(* IEC 61131-3 sources: 2026_Projet_YGO_ExcavatriceDragage/TOOLS/TEST_AUTO_CI/RESULTS/L_SIMULATION/tests (part 3) *)

(* ---- test_fb_sim_position_sensor.st ---- *)
(* T300 - Tests unitaires du capteur cumulatif M3. *)
TEST 'TC-T300-SEN-010 Hysteresis cumulative conserve le mot thermometre'
VAR
    fb : FB_Sim_PositionSensor;
END_VAR
    fb.Enable := TRUE;
    fb.Threshold_M := 5.0;
    fb.Hysteresis_M := 0.02;
    fb.Position_M := 4.99;
    fb();
    ASSERT_TRUE(fb.ElectricalOutput, 'Position sous seuil active DI cumulative');
    fb.Position_M := 5.01;
    fb();
    ASSERT_TRUE(fb.ElectricalOutput, 'Hysteresis maintient DI dans la bande');
    fb.Position_M := 5.03;
    fb();
    ASSERT_FALSE(fb.ElectricalOutput, 'Sortie au-dessus de seuil+hysteresis');
    fb.Position_M := 4.99;
    fb();
    ASSERT_FALSE(fb.ElectricalOutput, 'Retour dans bande ne re-declenche pas');
    fb.Position_M := 4.97;
    fb();
    ASSERT_TRUE(fb.ElectricalOutput, 'Retour sous seuil-hysteresis re-declenche');
END_TEST

TEST 'TC-T300-SEN-030 Episode intermittent est borne et rejoint la position'
VAR
    fb : FB_Sim_PositionSensor;
    i : INT;
END_VAR
    fb.Enable := TRUE;
    fb.Threshold_M := 5.0;
    fb.Position_M := 4.0;
    fb.IntermittenceActive := TRUE;
    fb.IntermittenceDurationS := 1.0;
    fb.IntermittencePeriodS := 0.12;
    fb.CycleTimeS := 0.01;
    fb();
    fb.Position_M := 6.0;
    FOR i := 1 TO 120 DO
        fb();
    END_FOR;
    ASSERT_FALSE(fb.EpisodeActive, 'Episode termine avant 1.2 s');
    ASSERT_FALSE(fb.ElectricalOutput, 'DI rejoint l etat mecanique final');
    ASSERT_GT(fb.TransitionCount, 2, 'Pertes/reprises publiees, sans front permanent');
END_TEST

TEST 'TC-T300-SEN-031 Recroisements mecaniques ne reinitialisent pas episode'
VAR
    fb : FB_Sim_PositionSensor;
    i : INT;
END_VAR
    fb.Enable := TRUE;
    fb.Threshold_M := 5.0;
    fb.Position_M := 4.0;
    fb.IntermittenceActive := TRUE;
    fb.IntermittenceDurationS := 1.0;
    fb.IntermittencePeriodS := 0.12;
    fb.CycleTimeS := 0.01;
    fb();
    FOR i := 1 TO 40 DO
        IF (i MOD 2) = 0 THEN
            fb.Position_M := 4.0;
        ELSE
            fb.Position_M := 6.0;
        END_IF;
        fb();
    END_FOR;
    fb.Position_M := 6.0;
    FOR i := 1 TO 70 DO
        fb();
    END_FOR;
    ASSERT_FALSE(fb.EpisodeActive, 'Recroisements ne prolongent pas episode au-dela de 1 s');
    ASSERT_FALSE(fb.ElectricalOutput, 'Etat final suit dernier franchissement mecanique');
END_TEST

TEST 'TC-T300-SEN-040 Cent graines deterministes bornent la stabilisation'
VAR
    fb : FB_Sim_PositionSensor;
    i : INT;
    j : INT;
END_VAR
    FOR i := 1 TO 100 DO
        fb.Enable := FALSE;
        fb();
        fb.Enable := TRUE;
        fb.Threshold_M := 5.0;
        fb.Position_M := 4.0;
        fb.IntermittenceActive := TRUE;
        fb.IntermittenceDurationS := 1.0;
        fb.IntermittencePeriodS := 0.12;
        fb.CycleTimeS := 0.01;
        fb.ScenarioSeed := DINT_TO_UDINT(i);
        fb();
        fb.Position_M := 6.0;
        FOR j := 1 TO 120 DO
            fb();
        END_FOR;
        ASSERT_FALSE(fb.EpisodeActive, 'Chaque graine termine son episode avant 1.2 s');
        ASSERT_FALSE(fb.ElectricalOutput, 'Chaque graine rejoint la position finale');
        ASSERT_GE(fb.EpisodeTogglePeriodS, 0.084, 'Periode aleatoire >= 70 % nominal');
        ASSERT_LE(fb.EpisodeTogglePeriodS, 0.156, 'Periode aleatoire <= 130 % nominal');
    END_FOR;
END_TEST

(* T300 P-A / C1-C2 — profil « BLIP COURT » : excursions electriques courtes, parametrables,
   independantes du train ~1 s ci-dessus. Signatures de la trace terrain du 2026-09-04 :
   Tremie contradictoire pendant 2 echantillons a 12,24 s ; PV reactive 1 echantillon a 14,94 s.
   Grille de test = 100 ms, celle de la trace. *)
TEST 'TC-T300-SEN-050 Blip court : largeur parametrable, deux sens, profil 1 s intact'
VAR
    fb : FB_Sim_PositionSensor;
    i : INT;
    excursions : INT;
    baseCount : UDINT;
END_VAR
    (* ---- (1) Sortie de zone, excursion 0,1 s => 1 echantillon (signature PV) ---- *)
    fb.Enable := TRUE;
    fb.Threshold_M := 5.0;
    fb.Hysteresis_M := 0.02;
    fb.CycleTimeS := 0.1;
    fb.ElectricalDelayS := 0.0;
    fb.Position_M := 4.0;
    fb();
    ASSERT_TRUE(fb.ElectricalOutput, 'Depart : dans la zone capteur');
    baseCount := fb.TransitionCount;
    fb.BlipTransitions := 1;
    fb.BlipDurationS := 0.1;
    fb.Position_M := 6.0;
    fb();
    excursions := 0;
    FOR i := 1 TO 6 DO
        fb();
        IF fb.ElectricalOutput <> fb.RawDetected THEN
            excursions := excursions + 1;
        END_IF;
    END_FOR;
    ASSERT_EQ(excursions, 1, 'Blip 0,1 s a 100 ms = 1 echantillon contradictoire');
    ASSERT_EQ(fb.TransitionCount - baseCount, 3, '1 front nominal + 2 fronts du blip');
    ASSERT_FALSE(fb.BlipActive, 'Blip borne et termine');
    ASSERT_FALSE(fb.ElectricalOutput, 'Sortie rendue a l etat mecanique final');

    (* ---- (2) Meme sens, excursion 0,2 s => 2 echantillons (signature Tremie) ---- *)
    fb.Enable := FALSE;
    fb();
    fb.Enable := TRUE;
    fb.BlipTransitions := 1;
    fb.BlipDurationS := 0.2;
    fb.Position_M := 4.0;
    fb();
    fb.Position_M := 6.0;
    fb();
    excursions := 0;
    FOR i := 1 TO 8 DO
        fb();
        IF fb.ElectricalOutput <> fb.RawDetected THEN
            excursions := excursions + 1;
        END_IF;
    END_FOR;
    ASSERT_EQ(excursions, 2, 'Blip 0,2 s a 100 ms = 2 echantillons contradictoires');
    ASSERT_FALSE(fb.ElectricalOutput, 'Sortie rendue a l etat mecanique final');

    (* ---- (3) Sens INVERSE : entree en zone (front montant) — symetrie AC5 ---- *)
    fb.Enable := FALSE;
    fb();
    fb.Enable := TRUE;
    fb.BlipTransitions := 1;
    fb.BlipDurationS := 0.2;
    fb.Position_M := 6.0;
    fb();
    ASSERT_FALSE(fb.ElectricalOutput, 'Depart : hors zone capteur');
    fb.Position_M := 4.0;
    fb();
    excursions := 0;
    FOR i := 1 TO 8 DO
        fb();
        IF fb.ElectricalOutput <> fb.RawDetected THEN
            excursions := excursions + 1;
        END_IF;
    END_FOR;
    ASSERT_EQ(excursions, 2, 'Symetrie : excursion equivalente a l entree en zone');
    ASSERT_TRUE(fb.ElectricalOutput, 'Sortie rendue a l etat mecanique final (dans la zone)');

    (* ---- (4) Blip DESACTIVE : le profil historique reste strictement inchange ---- *)
    fb.Enable := FALSE;
    fb();
    fb.Enable := TRUE;
    fb.BlipTransitions := 0;
    fb.Position_M := 4.0;
    fb();
    baseCount := fb.TransitionCount;
    fb.Position_M := 6.0;
    fb();
    excursions := 0;
    FOR i := 1 TO 10 DO
        fb();
        IF fb.ElectricalOutput <> fb.RawDetected THEN
            excursions := excursions + 1;
        END_IF;
    END_FOR;
    ASSERT_EQ(excursions, 0, 'Blip desactive : aucune excursion inventee');
    ASSERT_EQ(fb.TransitionCount - baseCount, 1, 'Blip desactive : seul le front nominal');
END_TEST

(* ---- test_fb_sim_safety.st ---- *)
(* =======================================================================
   Automated Unit Test - FB_Sim_Safety
   ======================================================================= *)
TEST 'TC-P13-SAF-001 Enable FALSE -> boucle AU ouverte'
VAR
    fb : FB_Sim_Safety;
END_VAR
    fb.Enable := FALSE;
    fb.SimChainOkBit := TRUE;
    fb();
    ASSERT_FALSE(fb.SimChainOk, 'Enable FALSE -> SimChainOk FALSE');
    ASSERT_FALSE(fb.SimContactorOk, 'Enable FALSE -> SimContactorOk FALSE');
END_TEST

TEST 'TC-P13-SAF-002 Pilotage boucle AU saine par SimChainOkBit et armement contacteur'
VAR
    fb : FB_Sim_Safety;
END_VAR
    fb.Enable := TRUE;
    fb.SimChainOkBit := TRUE; (* Chaine AU fermee par operateur *)
    fb();

    (* Ecoulement tempo de fermeture chaine (50ms = 60ms avancee) *)
    ADVANCE_TIME(60000000);
    fb();
    ASSERT_TRUE(fb.SimChainOk, 'SimChainOkBit TRUE -> SimChainOk TRUE apres tempo relais');

    (* Impulsion armement tenue 100ms (temps de collage contacteur) *)
    ADVANCE_TIME(10000000);
    fb.EmergencyArming := TRUE;
    fb();
    ADVANCE_TIME(110000000);
    fb();
    ASSERT_TRUE(fb.SimContactorOk, 'EmergencyArming soutenu -> SimContactorOk TRUE (engage)');

    (* Relachement impulsion -> auto-maintien *)
    ADVANCE_TIME(10000000);
    fb.EmergencyArming := FALSE;
    fb();
    ASSERT_TRUE(fb.SimContactorOk, 'Fin pulse -> Auto-maintien contacteur maintenu');
END_TEST

TEST 'TC-T306-SAF-003 Injection defaut rotation de phases par SimPhaseRotationOkBit'
VAR
    fb : FB_Sim_Safety;
END_VAR
    (* Phases saines : SimPhaseRotationOkBit=TRUE -> sortie TRUE (aucun defaut) *)
    fb.Enable := TRUE;
    fb.SimPhaseRotationOkBit := TRUE;
    fb();
    ASSERT_TRUE(fb.SimPhaseRotationOk, 'SimPhaseRotationOkBit TRUE -> SimPhaseRotationOk TRUE (phases saines)');

    (* Defaut injecte : SimPhaseRotationOkBit=FALSE -> sortie FALSE (PhaseRotationOk_DI tombe) *)
    fb.SimPhaseRotationOkBit := FALSE;
    fb();
    ASSERT_FALSE(fb.SimPhaseRotationOk, 'SimPhaseRotationOkBit FALSE -> SimPhaseRotationOk FALSE (defaut rotation de phases)');

    (* Retour a sain : nouveau passage a TRUE -> sortie TRUE *)
    fb.SimPhaseRotationOkBit := TRUE;
    fb();
    ASSERT_TRUE(fb.SimPhaseRotationOk, 'SimPhaseRotationOkBit TRUE apres FALSE -> SimPhaseRotationOk TRUE');
END_TEST

(* ---- test_fb_sim_suspended_load.st ---- *)
TEST 'TC-T300-MEC-010 Charge au repos ne cree pas d energie'
VAR
    fb : FB_Sim_SuspendedLoad;
    i : INT;
END_VAR
    fb.Enable := TRUE;
    fb.CycleTime_S := 0.01;
    FOR i := 1 TO 6000 DO
        fb();
    END_FOR;
    ASSERT_EQ(fb.Angle_Rad, 0.0, 'Angle nul sans excitation pendant 60 s');
    ASSERT_EQ(fb.AngularVelocity_RadPerS, 0.0, 'Vitesse angulaire nulle sans excitation');
END_TEST

TEST 'TC-T300-MEC-040 Acceleration excite charge et reaction reste conditionnee au frein'
VAR
    fb : FB_Sim_SuspendedLoad;
    i : INT;
END_VAR
    fb.Enable := TRUE;
    fb.CartAcceleration_Mps2 := 1.0;
    fb.BrakeMechanicallyOpen := FALSE;
    fb.CycleTime_S := 0.01;
    fb();
    ASSERT_TRUE(ABS(fb.Angle_Rad) > 0.0, 'Acceleration excite le pendule');
    ASSERT_EQ(fb.VelocityReaction_Mps, 0.0, 'Frein serre bloque reaction chariot');
    fb.BrakeMechanicallyOpen := TRUE;
    fb.CartAcceleration_Mps2 := 0.0;
    FOR i := 1 TO 10 DO
        fb();
    END_FOR;
    ASSERT_TRUE(ABS(fb.VelocityReaction_Mps) > 0.0, 'Frein ouvert publie reaction charge');
END_TEST

TEST 'TC-T300-MEC-020 Convergence pendule entre pas 10 ms et 5 ms'
VAR
    fb10 : FB_Sim_SuspendedLoad;
    fb5 : FB_Sim_SuspendedLoad;
    i : INT;
END_VAR
    fb10.Enable := TRUE;
    fb10.BrakeMechanicallyOpen := TRUE;
    fb10.CartAcceleration_Mps2 := 1.0;
    fb10.CycleTime_S := 0.01;
    fb5.Enable := TRUE;
    fb5.BrakeMechanicallyOpen := TRUE;
    fb5.CartAcceleration_Mps2 := 1.0;
    fb5.CycleTime_S := 0.005;
    fb10();
    fb5();
    fb5();
    fb10.CartAcceleration_Mps2 := 0.0;
    fb5.CartAcceleration_Mps2 := 0.0;
    FOR i := 1 TO 100 DO
        fb10();
        fb5();
        fb5();
    END_FOR;
    ASSERT_LT(ABS(fb10.Angle_Rad - fb5.Angle_Rad), 0.01,
        'Ecart angle inferieur a 10 mrad apres 1 s');
    ASSERT_LT(ABS(fb10.VelocityReaction_Mps - fb5.VelocityReaction_Mps), 0.001,
        'Ecart reaction inferieur a 1 mm/s apres 1 s');
END_TEST

(* ---- test_fb_sim_translation.st ---- *)
(* T300 - Tests du modele dynamique M3. *)
TEST 'TC-T300-TR-001 Etat sur desactive est P1 sans mouvement'
VAR
    fb : FB_Sim_Translation;
END_VAR
    fb.Enable := FALSE;
    fb();
    ASSERT_FALSE(fb.PosTremie, 'P1 ne doit pas annoncer Tremie');
    ASSERT_TRUE(fb.PosP1, 'Etat de repli deterministe sur P1');
    ASSERT_TRUE(fb.PosMaintenance, 'Mot thermometre P1 attendu');
    ASSERT_EQ(fb.ActualFrequency_Hz, 0.0, 'Frequence nulle');
    ASSERT_FALSE(fb.BrakeContactOpen, 'Frein ferme');
END_TEST

(* T301/L1 -- the isolated model receives geometry and gain.  The static G518
   check proves the PRG_02 -> SimBench wiring; these cases prove that those
   inputs are actually consumed by the simulated plant. *)
TEST 'TC-T301-SRC-001 Position P1 recue initialise le chariot sans geometrie locale'
VAR
    fb : FB_Sim_Translation;
END_VAR
    fb.PosTremie_M := 2.0;
    fb.PosPV_M := 3.0;
    fb.PosP2_M := 5.0;
    fb.PosP1_M := 7.0;
    fb.PosMaintenance_M := 11.0;
    fb.Enable := FALSE;
    fb();
    ASSERT_NEAR(fb.PositionTrue_M, 7.0, 0.0001,
        'Repli positionne le chariot sur PosP1_M recu');
    ASSERT_TRUE(fb.PosP1, 'Repli publie P1 apres initialisation sur la position recue');
END_TEST

TEST 'TC-T301-SRC-002 Gain recu convertit la frequence retournee en vitesse'
VAR
    fb : FB_Sim_Translation;
    i : INT;
END_VAR
    fb.PosTremie_M := 0.0;
    fb.PosPV_M := 10.0;
    fb.PosP2_M := 20.0;
    fb.PosP1_M := 30.0;
    fb.PosMaintenance_M := 40.0;
    fb.GainMetersPerHzSec := 0.03;
    fb.MaxFreq_Hz := 20.0;
    fb.Enable := FALSE;
    fb();
    fb.Enable := TRUE;
    fb.ReqTremie := TRUE;
    fb.SpeedTgt_Pct := 100.0;
    fb.BrakeReleaseCmd := TRUE;
    fb.BrakeOpenDelayS := 0.0;
    fb.LoadReactionGain_Mps2 := 0.0;
    FOR i := 1 TO 400 DO
        fb();
    END_FOR;
    ASSERT_NEAR(fb.ActualFrequency_Hz, 20.0, 0.05,
        'Frequence maximale recue appliquee');
    ASSERT_NEAR(fb.VelocityTrue_Mps, -0.6, 0.02,
        'Vitesse = sens x gain recu x frequence retournee');
END_TEST

TEST 'TC-T300-SEN-010 Les deux extremites publient les mots thermometres valides'
VAR
    fb : FB_Sim_Translation;
    i : INT;
END_VAR
    fb.Enable := FALSE;
    fb();
    fb.Enable := TRUE;
    fb.ReqTremie := TRUE;
    fb.SpeedTgt_Pct := 100.0;
    fb.BrakeReleaseCmd := TRUE;
    fb.BrakeOpenDelayS := 0.0;
    fb.FullTravelTimeS := 0.5;
    fb.SensorElectricalDelayS := 0.0;
    FOR i := 1 TO 400 DO
        fb();
    END_FOR;
    ASSERT_TRUE(fb.PosTremie, 'Tremie active a la butee 0 m');
    ASSERT_TRUE(fb.PosPV, 'PV cumulatif actif a Tremie');
    ASSERT_TRUE(fb.PosP2, 'P2 cumulatif actif a Tremie');
    ASSERT_TRUE(fb.PosP1, 'P1 cumulatif actif a Tremie');
    ASSERT_TRUE(fb.PosMaintenance, 'Maintenance cumulatif actif a Tremie');
    ASSERT_EQ(fb.VelocityTrue_Mps, 0.0, 'Butee Tremie absorbe la vitesse chariot');

    fb.Enable := FALSE;
    fb();
    fb.Enable := TRUE;
    fb.ReqTremie := FALSE;
    fb.ReqMaintenance := TRUE;
    fb.SpeedTgt_Pct := 100.0;
    fb.BrakeReleaseCmd := TRUE;
    fb.BrakeOpenDelayS := 0.0;
    fb.FullTravelTimeS := 0.5;
    fb.SensorElectricalDelayS := 0.0;
    FOR i := 1 TO 400 DO
        fb();
    END_FOR;
    ASSERT_FALSE(fb.PosTremie, 'Tremie inactif a Maintenance');
    ASSERT_FALSE(fb.PosPV, 'PV inactif a Maintenance');
    ASSERT_FALSE(fb.PosP2, 'P2 inactif a Maintenance');
    ASSERT_FALSE(fb.PosP1, 'P1 inactif a Maintenance');
    ASSERT_FALSE(fb.PosMaintenance, 'Maintenance inactif a la butee pour mot 00000');
    ASSERT_EQ(fb.VelocityTrue_Mps, 0.0, 'Butee Maintenance absorbe la vitesse chariot');
END_TEST

TEST 'TC-T300-SEN-011 Le capteur PV commute au franchissement vers Tremie'
VAR
    fb : FB_Sim_Translation;
    i : INT;
    pvWasFalse : BOOL;
    pvTurnedTrue : BOOL;
END_VAR
    fb.Enable := TRUE;
    fb.ReqTremie := TRUE;
    fb.SpeedTgt_Pct := 100.0;
    fb.BrakeReleaseCmd := TRUE;
    fb.FullTravelTimeS := 8.0;
    fb.SensorElectricalDelayS := 0.0;
    pvWasFalse := FALSE;
    pvTurnedTrue := FALSE;
    FOR i := 1 TO 700 DO
        fb();
        IF NOT fb.PosPV THEN
            pvWasFalse := TRUE;
        END_IF;
        IF pvWasFalse AND fb.PosPV THEN
            pvTurnedTrue := TRUE;
        END_IF;
    END_FOR;
    ASSERT_TRUE(pvWasFalse, 'PV initialement inactif a P1');
    ASSERT_TRUE(pvTurnedTrue, 'PV actif apres franchissement vers Tremie');
END_TEST

TEST 'TC-T300-DRV-020 Rampe terrain 20 Hz par seconde'
VAR
    fb : FB_Sim_Translation;
    i : INT;
END_VAR
    fb.Enable := TRUE;
    fb.ReqTremie := TRUE;
    fb.SpeedTgt_Pct := 0.0;
    fb.BrakeReleaseCmd := TRUE;
    fb();
    fb.SpeedTgt_Pct := 100.0;
    FOR i := 1 TO 100 DO
        fb();
    END_FOR;
    ASSERT_GT(fb.FrequencyCmd_Hz, 19.7, 'Rampe apres 1 s >= 19.7 Hz');
    ASSERT_LT(fb.FrequencyCmd_Hz, 20.3, 'Rampe apres 1 s <= 20.3 Hz');
    ASSERT_LT(fb.ActualFrequency_Hz, fb.FrequencyCmd_Hz, 'Retour dynamique derriere la consigne');
    ASSERT_GT(fb.ActualFrequency_Hz, 16.0, 'Retour coherent avec tau 150 ms');
END_TEST

TEST 'TC-T300-BRK-025 Frein temporise et retour distinct'
VAR
    fb : FB_Sim_Translation;
    i : INT;
END_VAR
    fb.Enable := TRUE;
    fb.BrakeReleaseCmd := TRUE;
    fb.BrakeOpenDelayS := 0.10;
    fb();
    ASSERT_TRUE(fb.BrakeCoilEnergized, 'Bobine active immediatement sur ordre');
    FOR i := 1 TO 8 DO
        fb();
    END_FOR;
    ASSERT_FALSE(fb.BrakeContactOpen, 'Pas de confirmation avant 90 ms');
    fb();
    fb();
    ASSERT_TRUE(fb.BrakeMechanicallyOpen, 'Ouverture mecanique apres delai');
    ASSERT_TRUE(fb.BrakeContactOpen, 'Retour auxiliaire apres delai');
END_TEST

TEST 'TC-T300-MEC-010 Le chariot suit la frequence et excite la charge'
VAR
    fb : FB_Sim_Translation;
    i : INT;
    startPosition_M : REAL;
END_VAR
    fb.Enable := TRUE;
    fb.ReqTremie := TRUE;
    fb.SpeedTgt_Pct := 100.0;
    fb.BrakeReleaseCmd := TRUE;
    fb.BrakeOpenDelayS := 0.0;
    fb();
    startPosition_M := fb.PositionTrue_M;
    FOR i := 1 TO 100 DO
        fb();
    END_FOR;
    ASSERT_LT(fb.PositionTrue_M, startPosition_M, 'Deplacement reel vers Tremie');
    ASSERT_LT(fb.VelocityTrue_Mps, 0.0, 'Vitesse signee vers Tremie');
    ASSERT_TRUE(ABS(fb.LoadAngle_Rad) > 0.0001, 'Acceleration excite le pendule');
END_TEST

TEST 'TC-T300-MEC-030 Commandes contradictoires restent neutres'
VAR
    fb : FB_Sim_Translation;
    i : INT;
    startPosition_M : REAL;
END_VAR
    fb.Enable := TRUE;
    fb.ReqTremie := TRUE;
    fb.ReqMaintenance := TRUE;
    fb.SpeedTgt_Pct := 100.0;
    fb.BrakeReleaseCmd := TRUE;
    fb.BrakeOpenDelayS := 0.0;
    fb();
    startPosition_M := fb.PositionTrue_M;
    FOR i := 1 TO 50 DO
        fb();
    END_FOR;
    ASSERT_EQ(fb.FrequencyCmd_Hz, 0.0, 'Aucune excitation avec deux sens');
    ASSERT_EQ(fb.PositionTrue_M, startPosition_M, 'Position conservee');
END_TEST

TEST 'TC-T300-SEN-030 Episode capteur intermittent rejouable avant stabilisation'
VAR
    fb : FB_Sim_Translation;
    i : INT;
END_VAR
    fb.Enable := TRUE;
    fb.ReqMaintenance := TRUE;
    fb.SpeedTgt_Pct := 0.0;
    fb.BrakeReleaseCmd := TRUE;
    fb.BrakeOpenDelayS := 0.0;
    fb.FullTravelTimeS := 0.5;
    fb.SensorStabilizationS := 1.0;
    fb.SensorIntermittenceActive := TRUE;
    fb.SensorLoadAngleTriggerRad := 0.0;
    fb.SensorIntermittencePeriodS := 0.12;
    fb();
    fb.SpeedTgt_Pct := 100.0;
    FOR i := 1 TO 250 DO
        fb();
    END_FOR;
    ASSERT_GT(fb.SensorTransitionCount, 1, 'Au moins deux fronts DI sont publies pendant episode');
    ASSERT_FALSE(fb.PosP1, 'DI rejoint la position mecanique apres episode');
END_TEST

TEST 'TC-T300-CAM-100 Matrice 48 scenarios par 100 graines respecte invariants'
VAR
    fb : FB_Sim_Translation;
    direction : INT;
    loadProfile : INT;
    regime : INT;
    perturbation : INT;
    seed : INT;
    i : INT;
END_VAR
    FOR direction := 1 TO 2 DO
        FOR loadProfile := 1 TO 2 DO
            FOR regime := 1 TO 3 DO
                FOR perturbation := 1 TO 4 DO
                    FOR seed := 1 TO 100 DO
                        fb.Enable := FALSE;
                        fb();
                        fb.Enable := TRUE;
                        fb.ReqTremie := direction = 1;
                        fb.ReqMaintenance := direction = 2;
                        fb.SpeedTgt_Pct := 100.0;
                        fb.BrakeReleaseCmd := TRUE;
                        fb.FullTravelTimeS := 0.5;
                        fb.SensorElectricalDelayS := 0.0;
                        fb.SensorScenarioSeed := DINT_TO_UDINT(seed);
                        fb.SensorIntermittenceActive := perturbation = 3;
                        fb.SensorLoadAngleTriggerRad := 0.0;
                        IF loadProfile = 1 THEN
                            fb.LoadReactionGain_Mps2 := 0.0;
                        ELSE
                            fb.LoadReactionGain_Mps2 := 0.20;
                        END_IF;
                        IF perturbation = 4 THEN
                            fb.BrakeOpenDelayS := 0.30;
                        ELSE
                            fb.BrakeOpenDelayS := 0.0;
                        END_IF;
                        fb();
                        FOR i := 1 TO 200 DO
                            IF (regime = 2) AND (i = 80) THEN
                                fb.SpeedTgt_Pct := 0.0;
                            ELSIF (regime = 3) AND (i = 80) THEN
                                fb.SpeedTgt_Pct := 0.0;
                                fb.BrakeReleaseCmd := FALSE;
                            END_IF;
                            fb();
                            ASSERT_GE(fb.PositionTrue_M, 0.0, 'Course mecanique jamais inferieure a Tremie');
                            ASSERT_LE(fb.PositionTrue_M, 30.0, 'Course mecanique jamais superieure a Maintenance');
                            ASSERT_GE(fb.ActualFrequency_Hz, 0.0, 'Retour variateur non negatif');
                            ASSERT_LE(fb.ActualFrequency_Hz, 50.0, 'Retour variateur borne a 50 Hz');
                            IF perturbation <> 3 THEN
                                ASSERT_TRUE((NOT fb.PosTremie) OR fb.PosPV,
                                    'Mot thermometre : Tremie implique PV');
                                ASSERT_TRUE((NOT fb.PosPV) OR fb.PosP2,
                                    'Mot thermometre : PV implique P2');
                                ASSERT_TRUE((NOT fb.PosP2) OR fb.PosP1,
                                    'Mot thermometre : P2 implique P1');
                                ASSERT_TRUE((NOT fb.PosP1) OR fb.PosMaintenance,
                                    'Mot thermometre : P1 implique Maintenance');
                            END_IF;
                        END_FOR;
                    END_FOR;
                END_FOR;
            END_FOR;
        END_FOR;
    END_FOR;
END_TEST

(* T300 P-A / C4 — traversee de la faute frein dans le composite : prouve que l'entree
   descend jusqu'a FB_Sim_TranslationBrake et que la sortie remonte, sans toucher au
   nominal (premier palier d'assertions). *)
TEST 'TC-T300-BRK-041 Faute frein traverse le composite M3 (fermeture en mouvement)'
VAR
    fb : FB_Sim_Translation;
    i : INT;
END_VAR
    fb.Enable := TRUE;
    fb.ReqMaintenance := TRUE;
    fb.SpeedTgt_Pct := 100.0;
    fb.BrakeReleaseCmd := TRUE;
    fb.BrakeOpenDelayS := 0.0;
    fb();
    ASSERT_TRUE(fb.BrakeMechanicallyOpen, 'Frein ouvert au depart');
    FOR i := 1 TO 200 DO
        fb();
    END_FOR;
    ASSERT_GT(fb.ActualFrequency_Hz, 0.5, 'Chariot en mouvement (frequence non nulle)');
    ASSERT_TRUE(fb.BrakeMechanicallyOpen, 'NOMINAL : frein ouvert tant que la vitesse est non nulle');
    ASSERT_FALSE(fb.BrakeFaultCloseActive, 'Aucune faute par defaut');

    fb.BrakeFaultCloseWhileRunning := TRUE;
    FOR i := 1 TO 12 DO
        fb();
    END_FOR;
    ASSERT_TRUE(fb.BrakeFaultCloseActive, 'Faute frein relayee par le composite');
    ASSERT_GT(fb.ActualFrequency_Hz, 0.5, 'Vitesse encore non nulle a la fermeture');
    ASSERT_FALSE(fb.BrakeMechanicallyOpen, 'Faute : frein mecaniquement serre en mouvement');
END_TEST

(* T300 P-A / C3 — deceleration libre. Trace terrain 2026-09-04 : commande retiree a
   14,67 s alors que 33,98 Hz etaient retournes ; le chariot a continue d'avancer pendant
   1,49 s jusqu'a l'arret a 16,16 s. La distance de roue libre correspondante est une
   ESTIMATION (la trace ne contient aucune variable de position) : ordre de grandeur
   1,1 a 1,3 m selon la methode d'integration, jamais parcourus par le modele avant ce
   correctif qui annulait la vitesse au scan de retrait de commande.
   Le pas FullTravelTimeS est allonge (60 s) pour que le scenario reste loin des butees
   mecaniques et que l'oracle porte sur la SEULE deceleration libre, pas sur un choc. *)
TEST 'TC-T300-DRV-070 Deceleration libre : le chariot avance encore apres retrait de commande'
VAR
    fb : FB_Sim_Translation;
    i : INT;
    posAtCut_M : REAL;
END_VAR
    fb.Enable := TRUE;
    fb.ReqMaintenance := TRUE;
    fb.SpeedTgt_Pct := 100.0;
    fb.BrakeReleaseCmd := TRUE;
    fb.BrakeOpenDelayS := 0.0;
    (* Echelle par defaut du banc : palier 50 Hz (maximum variateur), 0,02 m/(Hz.s), rampe d'arret 25 Hz/s. *)
    (* Charge neutralisee : l'oracle porte sur la SEULE deceleration libre du variateur.
       Sans cela, le droop de charge (0,5 Hz par rad/s) peut faire passer ActualFrequency
       sous 39,5 Hz et rendre l'assertion de palier marginale — bruit, pas verite. *)
    fb.LoadFrequencyDroopGain_Hz := 0.0;
    fb.LoadReactionGain_Mps2 := 0.0;
    FOR i := 1 TO 400 DO
        fb();
    END_FOR;
    ASSERT_NEAR(fb.ActualFrequency_Hz, 50.0, 0.5, 'Palier 50 Hz etabli avant le retrait');
    ASSERT_LT(fb.PositionTrue_M, 30.0, 'Chariot encore hors butee (scenario non pollue)');

    (* Retrait total de la commande : plus aucune requete, consigne a zero. *)
    fb.ReqMaintenance := FALSE;
    fb.ReqTremie := FALSE;
    fb.SpeedTgt_Pct := 0.0;
    fb();
    ASSERT_GT(fb.ActualFrequency_Hz, 0.5, 'Le variateur retourne encore de la vitesse au retrait');
    posAtCut_M := fb.PositionTrue_M;

    (* Roue libre : la position doit continuer de varier tant que ActualFrequency_Hz > 0.
       Seuil = borne BASSE de la bande de reference trace (R2-O9 : 0,9 a 1,3 m). Le modele
       parcourt davantage (~2,2 m) car sa rampe de descente dure 2,0 s contre 1,49 s mesures :
       ecart de fidelite ASSUME, borne haute verifiee separement. Avant correctif : ~0,1 m. *)
    FOR i := 1 TO 300 DO
        fb();
    END_FOR;
    ASSERT_NEAR(fb.ActualFrequency_Hz, 0.0, 0.01, 'Retour variateur revenu a zero');
    ASSERT_GE(fb.PositionTrue_M - posAtCut_M, 0.9,
        'Roue libre >= borne basse trace (avant correctif : ~0,1 m)');
    ASSERT_LE(fb.PositionTrue_M - posAtCut_M, 3.0, 'Roue libre bornee (pas d emballement)');
    ASSERT_LE(fb.PositionTrue_M, 30.0, 'Course mecanique respectee');
END_TEST

(* T300 P-A / C5 — perte DEFINITIVE du capteur Tremie apres arret serre.
   Trace terrain 2026-09-04 : a 26,437 s le chariot entre en zone Tremie pendant que la
   commande est retiree ; le capteur retombe a 26,537 s et n'est JAMAIS repris sur les
   8,6 s restantes (PLAN_T300 §38 : perte unique post-arret, pas une oscillation entretenue).
   EndStopRecoilMax_M = 0 conserve le comportement historique (position ET vitesse figees,
   decision de review tracee) : les deux regimes sont verifies ici. *)
TEST 'TC-T300-SEN-052 Recul borne a la butee Tremie : DI perdue PUIS reprise oscillante (ecart trace)'
VAR
    fb : FB_Sim_Translation;
    i : INT;
    scansToFall : INT;
    scansActive : INT;
END_VAR
    (* --- (0) NON-REGRESSION : recul non autorise => comportement historique inchange --- *)
    fb.Enable := TRUE;
    fb.ReqTremie := TRUE;
    fb.SpeedTgt_Pct := 100.0;
    fb.BrakeReleaseCmd := TRUE;
    fb.BrakeOpenDelayS := 0.0;
    fb.SensorElectricalDelayS := 0.0;
    fb.EndStopRecoilMax_M := 0.0;
    (* T361 — pas de temps PINCE ici : l'oracle de ce cas est le recul a la butee, pas
       l'echelle odometrique. Le scenario vient de la trace du 2026-09-04 (quelques
       secondes de trajet) et le defaut du FB est passe de 8,0 s a 37,5 s pour s'aligner
       sur le gain reel : sans ce pas explicite, 900 scans (9 s) ne suffiraient plus a
       atteindre la butee Tremie depuis 20 m et le cas testerait autre chose que son objet. *)
    fb.FullTravelTimeS := 8.0;
    FOR i := 1 TO 900 DO
        fb();
    END_FOR;
    ASSERT_TRUE(fb.PosTremie, 'Historique : DI Tremie TENUE a la butee quand le recul est interdit');
    ASSERT_NEAR(fb.PositionTrue_M, 0.0, 0.001, 'Historique : position figee a la butee');

    (* --- (1) Recul borne autorise : la charge ressort le chariot de la zone --- *)
    fb.Enable := FALSE;
    fb();
    fb.Enable := TRUE;
    fb.EndStopRecoilMax_M := 0.5;
    fb.LoadReactionGain_Mps2 := 2.0;
    FOR i := 1 TO 900 DO
        fb();
    END_FOR;
    ASSERT_TRUE(fb.PosTremie, 'PRECONDITION : zone Tremie atteinte (recul = 0,5 m autorise)');

    (* Commande retiree a l'instant de l' entree en zone (sequence exacte de la trace). *)
    fb.ReqTremie := FALSE;
    fb.SpeedTgt_Pct := 0.0;
    scansToFall := 0;
    FOR i := 1 TO 600 DO
        fb();
        IF (NOT fb.PosTremie) AND (scansToFall = 0) THEN
            scansToFall := i;
        END_IF;
    END_FOR;
    ASSERT_GT(scansToFall, 0, 'DI Tremie RETOMBE apres l arret serre (recul borne)');
    (* Boucle a 600 scans, seuil a 300 : assertion NON tautologique, marge reelle au-dessus
       de la valeur mesuree (256 scans). *)
    ASSERT_LE(scansToFall, 300, 'Perte dans un temps borne (<= 3 s a 10 ms)');

    (* Perte DURABLE : le capteur ne se reactive pas de facon entretenue ensuite. *)
    scansActive := 0;
    FOR i := 1 TO 500 DO
        fb();
        IF fb.PosTremie THEN
            scansActive := scansActive + 1;
        END_IF;
    END_FOR;
    (* ⚠️ LIMITE CONNUE — NON MASQUEE. Le modele reduit n'a AUCUNE friction de chariot ni
       raideur de cable : le pendule amorti ramene le chariot dans la zone capteur par
       oscillations. La perte est donc BORNEE, mais pas encore DEFINITIVE comme sur la trace
       terrain (PLAN_T300 §38 : « perte unique post-arret, pas une oscillation entretenue »).
       Fermer cet ecart exige un parametre physique nouveau (friction de roulement / raideur
       de cable), hors perimetre de ce lot et non calibrable sans mesure terrain : ce test
       CARACTERISE l'etat reel, il ne le valide pas. Mesure : 106 scans actifs sur 500
       (21 %), contre 0 attendu par la trace. Assertion volontairement en enveloppe. *)
    ASSERT_LE(scansActive, 150, 'Perte BORNEE mais NON DEFINITIVE : ecart trace documente');
END_TEST

(* =========================================================================
   T361 VOLET A — ALIGNEMENT DU RATIO ODOMETRIQUE BANC / ESTIMATEUR
   =========================================================================
   Le banc et l'estimateur integrent la MEME frequence retournee, mais avec deux
   echelles construites separement :
     - estimateur (CODE/I_TRANSLATION/FB_Translation_PositionEstimator.st:153/155) :
       dx = f x GainMetersPerHzSec x dt, gain cable en PRG_05_Translation.st:591 sur
       GVL_PERSISTENT._TranslationGainMetersPerHzSec = 0,02 m/(Hz.s) (1 m/s a 50 Hz) ;
     - banc (ce FB) : dx = f x (CST_PositionAtMaintenance / (40 x FullTravelTimeS)) x dt.
   Tant que les deux echelles divergent, la position estimee prend un retard constant et
   CHAQUE franchissement de capteur produit un saut de recalage — c'est exactement ce que
   montre la trace Suivi_74 (sauts de 4,53 / 9,12 / 4,59 m, AUDIT_T360). Avec l'echelle
   historique 8,0 s le rapport valait 0,09375 / 0,02 = 4,7.
   Les deux cas ci-dessous comparent le banc a l'expression EXACTE de l'estimateur :
   ils echouent si l'une des deux echelles bouge sans l'autre. *)

TEST 'TC-T361-ALIGN-001 Ratio odometrique du banc = gain reel 0,02 m/(Hz.s)'
VAR
    fb : FB_Sim_Translation;
    i : INT;
END_VAR
    fb.Enable := TRUE;
    fb.ReqMaintenance := TRUE;
    fb.SpeedTgt_Pct := 100.0;
    fb.BrakeReleaseCmd := TRUE;
    fb.BrakeOpenDelayS := 0.0;
    (* Charge neutralisee : l'oracle porte sur l'ECHELLE seule, pas sur la reaction du pendule. *)
    fb.LoadReactionGain_Mps2 := 0.0;
    FOR i := 1 TO 400 DO
        fb();
    END_FOR;
    ASSERT_NEAR(fb.ActualFrequency_Hz, 50.0, 0.5, 'Palier 50 Hz (maximum variateur) etabli avant lecture du ratio');
    ASSERT_NEAR(fb.VelocityTrue_Mps / fb.ActualFrequency_Hz, 0.02, 0.0002,
        'Ratio banc (m/s par Hz) = _TranslationGainMetersPerHzSec (ancien : 0,09375)');
END_TEST

TEST 'TC-T361-ALIGN-002 Distance banc = integrale f x 0,02 m/(Hz.s) sur 6 s'
VAR
    fb : FB_Sim_Translation;
    i : INT;
    posStart_M : REAL;
    integralHzS : REAL;
END_VAR
    fb.Enable := TRUE;
    fb.ReqTremie := TRUE;
    fb.SpeedTgt_Pct := 100.0;
    fb.BrakeReleaseCmd := TRUE;
    fb.BrakeOpenDelayS := 0.0;
    fb.SensorElectricalDelayS := 0.0;
    fb.LoadReactionGain_Mps2 := 0.0;
    (* 2 s pour etablir le palier, puis 6 s de mesure (600 scans a 10 ms) largement
       a l'ecart des butees : 20 m -> ~15,2 m a 0,8 m/s. *)
    FOR i := 1 TO 200 DO
        fb();
    END_FOR;
    posStart_M := fb.PositionTrue_M;
    integralHzS := 0.0;
    FOR i := 1 TO 600 DO
        fb();
        integralHzS := integralHzS + fb.ActualFrequency_Hz * 0.010;
    END_FOR;
    (* Tolerance 0,25 m (soit ~5 % de 4,8 m) : elle couvre la seule trainee de 1er ordre du
       modele de vitesse, pas une erreur d'echelle — un ecart d'echelle de 4,7 ferait
       diverger les deux membres de plusieurs metres. *)
    ASSERT_NEAR(posStart_M - fb.PositionTrue_M, integralHzS * 0.02, 0.25,
        'Distance parcourue par le banc = position reconstituee par l estimateur odometrique');
END_TEST

(* Echelle de la consigne : PRG_02 envoie SpeedCmd_Pct = f / 50 Hz x 100.
   20 Hz d'approche reels = 40 % doivent redonner 20 Hz (pas 16 Hz). Charge neutralisee. *)
TEST 'TC-T417-SCALE-001 Consigne 40 pct = 20 Hz et 100 pct = 50 Hz'
VAR
    fbApproach : FB_Sim_Translation;
    fbMax : FB_Sim_Translation;
    i : INT;
END_VAR
    fbApproach.Enable := TRUE;
    fbApproach.ReqMaintenance := TRUE;
    fbApproach.SpeedTgt_Pct := 40.0;
    fbApproach.BrakeReleaseCmd := TRUE;
    fbApproach.BrakeOpenDelayS := 0.0;
    fbApproach.LoadFrequencyDroopGain_Hz := 0.0;
    fbApproach.LoadReactionGain_Mps2 := 0.0;
    fbMax.Enable := TRUE;
    fbMax.ReqMaintenance := TRUE;
    fbMax.SpeedTgt_Pct := 100.0;
    fbMax.BrakeReleaseCmd := TRUE;
    fbMax.BrakeOpenDelayS := 0.0;
    fbMax.LoadFrequencyDroopGain_Hz := 0.0;
    fbMax.LoadReactionGain_Mps2 := 0.0;
    FOR i := 1 TO 400 DO
        fbApproach();
        fbMax();
    END_FOR;
    ASSERT_NEAR(fbApproach.ActualFrequency_Hz, 20.0, 0.05, '40 pct de 50 Hz = 20 Hz en regime etabli');
    ASSERT_NEAR(fbMax.ActualFrequency_Hz, 50.0, 0.05, '100 pct = 50 Hz (maximum variateur)');
END_TEST

(* Rampe d'arret : trace reelle ~25 Hz/s (rampe variateur). Pente mesuree sur la fenetre
   utile 10 Hz -> ~4 Hz, apres le transitoire du filtre de 1er ordre. Charge neutralisee. *)
TEST 'TC-T417-DECEL-001 Pente d arret 25 Hz/s depuis l approche 20 Hz'
VAR
    fb : FB_Sim_Translation;
    i : INT;
    f1_Hz : REAL;
END_VAR
    fb.Enable := TRUE;
    fb.ReqMaintenance := TRUE;
    fb.SpeedTgt_Pct := 40.0;
    fb.BrakeReleaseCmd := TRUE;
    fb.BrakeOpenDelayS := 0.0;
    fb.LoadFrequencyDroopGain_Hz := 0.0;
    fb.LoadReactionGain_Mps2 := 0.0;
    FOR i := 1 TO 400 DO
        fb();
    END_FOR;
    ASSERT_NEAR(fb.ActualFrequency_Hz, 20.0, 0.05, 'Approche 20 Hz etablie avant le retrait');
    fb.SpeedTgt_Pct := 0.0;
    i := 0;
    WHILE (fb.ActualFrequency_Hz > 10.0) AND (i < 300) DO
        fb();
        i := i + 1;
    END_WHILE;
    f1_Hz := fb.ActualFrequency_Hz;
    FOR i := 1 TO 20 DO
        fb();
    END_FOR;
    ASSERT_NEAR((f1_Hz - fb.ActualFrequency_Hz) / 0.2, 25.0, 1.0, 'Pente de decroissance = 25 Hz/s');
END_TEST

(* Depassement apres retrait de commande a l'approche : ordre de grandeur de la trace reelle
   (~0,25 m, gain 0,02 m/(Hz.s) provisoire). Bande large : cible a confirmer par la trace 10 ms. *)
TEST 'TC-T417-OVERSHOOT-001 Depassement apres retrait a 20 Hz'
VAR
    fb : FB_Sim_Translation;
    i : INT;
    posAtCut_M : REAL;
    overshoot_M : REAL;
END_VAR
    fb.Enable := TRUE;
    fb.ReqMaintenance := TRUE;
    fb.SpeedTgt_Pct := 40.0;
    fb.BrakeReleaseCmd := TRUE;
    fb.BrakeOpenDelayS := 0.0;
    fb.LoadFrequencyDroopGain_Hz := 0.0;
    fb.LoadReactionGain_Mps2 := 0.0;
    FOR i := 1 TO 400 DO
        fb();
    END_FOR;
    ASSERT_NEAR(fb.ActualFrequency_Hz, 20.0, 0.05, 'Approche 20 Hz etablie avant le retrait');
    fb.ReqMaintenance := FALSE;
    fb.SpeedTgt_Pct := 0.0;
    fb();
    posAtCut_M := fb.PositionTrue_M;
    FOR i := 1 TO 300 DO
        fb();
    END_FOR;
    overshoot_M := fb.PositionTrue_M - posAtCut_M;
    ASSERT_GE(overshoot_M, 0.15, 'Depassement >= 0,15 m (ordre de grandeur trace reelle)');
    ASSERT_LE(overshoot_M, 0.35, 'Depassement <= 0,35 m (ordre de grandeur trace reelle)');
END_TEST

(* Acceleration du banc : chariot ET frequence retournee x facteur. L'estimateur reel integre
   f_retournee x 0,02 : il doit retrouver la distance du chariot (aucun saut de recalage). *)
TEST 'TC-SIMSPEED-001 Facteur 3 : chariot 3 m/s a 50 Hz et distance = integrale f retournee x 0,02'
VAR
    fb : FB_Sim_Translation;
    i : INT;
    posStart_M : REAL;
    integralHzS : REAL;
END_VAR
    fb.Enable := TRUE;
    fb.ReqTremie := TRUE;
    fb.SpeedTgt_Pct := 100.0;
    fb.SpeedFactor := 3.0;
    fb.BrakeReleaseCmd := TRUE;
    fb.BrakeOpenDelayS := 0.0;
    fb.SensorElectricalDelayS := 0.0;
    fb.LoadReactionGain_Mps2 := 0.0;
    FOR i := 1 TO 300 DO
        fb();
    END_FOR;
    ASSERT_NEAR(fb.ActualFrequency_Hz, 150.0, 3.0, 'frequence retournee = 3 x 50 Hz');
    ASSERT_NEAR(fb.VelocityTrue_Mps, -3.0, 0.15, 'chariot a 3 m/s (1 m/s reel x 3)');
    posStart_M := fb.PositionTrue_M;
    integralHzS := 0.0;
    FOR i := 1 TO 200 DO
        fb();
        integralHzS := integralHzS + fb.ActualFrequency_Hz * 0.010;
    END_FOR;
    ASSERT_NEAR(posStart_M - fb.PositionTrue_M, integralHzS * 0.02, 0.25,
        'estimation (f retournee x 0,02) = distance du chariot : aucun saut de recalage');
END_TEST

TEST 'TC-SIMSPEED-002 Facteur borne a 5, facteur < 1 ramene a 1'
VAR
    fb : FB_Sim_Translation;
    fbLow : FB_Sim_Translation;
    i : INT;
END_VAR
    fb.Enable := TRUE;
    fb.ReqTremie := TRUE;
    fb.SpeedTgt_Pct := 100.0;
    fb.SpeedFactor := 10.0;
    fb.BrakeReleaseCmd := TRUE;
    fb.BrakeOpenDelayS := 0.0;
    fb.LoadReactionGain_Mps2 := 0.0;
    fbLow.Enable := TRUE;
    fbLow.ReqTremie := TRUE;
    fbLow.SpeedTgt_Pct := 100.0;
    fbLow.SpeedFactor := 0.0;
    fbLow.BrakeReleaseCmd := TRUE;
    fbLow.BrakeOpenDelayS := 0.0;
    fbLow.LoadReactionGain_Mps2 := 0.0;
    FOR i := 1 TO 300 DO
        fb();
        fbLow();
    END_FOR;
    ASSERT_NEAR(fb.ActualFrequency_Hz, 250.0, 5.0, 'facteur 10 borne a 5 : 250 Hz retournes');
    ASSERT_NEAR(fbLow.ActualFrequency_Hz, 50.0, 1.0, 'facteur 0 ramene a 1 : 50 Hz retournes');
    ASSERT_NEAR(fbLow.VelocityTrue_Mps, -1.0, 0.05, 'facteur 1 : 1 m/s reel a 50 Hz');
END_TEST

(* ---- test_fb_sim_translation_brake.st ---- *)
TEST 'TC-T300-BRK-010 Bobine mecanique et contact restent distincts'
VAR
    fb : FB_Sim_TranslationBrake;
    i : INT;
END_VAR
    fb.Enable := TRUE;
    fb.ReleaseCmd := TRUE;
    fb.OpenDelay_S := 0.10;
    fb.ContactDelay_S := 0.01;
    fb.CycleTime_S := 0.01;
    FOR i := 1 TO 9 DO
        fb();
    END_FOR;
    ASSERT_TRUE(fb.CoilEnergized, 'Bobine immediate');
    ASSERT_FALSE(fb.MechanicallyOpen, 'Effet mecanique pas avant delai');
    fb();
    fb();
    ASSERT_TRUE(fb.MechanicallyOpen, 'Ouverture mecanique apres 100 ms');
    fb();
    ASSERT_TRUE(fb.ContactOpen, 'Contact apres effet mecanique');
END_TEST

TEST 'TC-T300-BRK-020 Serrage attend vitesse nulle'
VAR
    fb : FB_Sim_TranslationBrake;
    i : INT;
END_VAR
    fb.Enable := TRUE;
    fb.ReleaseCmd := TRUE;
    fb.OpenDelay_S := 0.0;
    fb.CycleTime_S := 0.01;
    fb();
    fb.ReleaseCmd := FALSE;
    fb.ActualFrequency_Hz := 2.0;
    FOR i := 1 TO 20 DO
        fb();
    END_FOR;
    ASSERT_TRUE(fb.MechanicallyOpen, 'Frein reste ouvert tant que vitesse non nulle');
    fb.ActualFrequency_Hz := 0.0;
    FOR i := 1 TO 10 DO
        fb();
    END_FOR;
    ASSERT_FALSE(fb.MechanicallyOpen, 'Frein serre apres 90 ms a vitesse nulle');
END_TEST

(* T300 P-A / C4 — rejeu EXACT du defaut terrain du 2026-09-04 (trace M3, 26,437 s) :
   contact frein ferme alors que le variateur retourne encore 10,00 Hz (State.ErrorId=64).
   La branche de FAUTE est explicite et le defaut de l'entree est FALSE : le chemin nominal
   reste celui de TC-T300-BRK-020, dont la garde 0,5 Hz est validee par la MEME trace
   (frein ouvert a 0,60 Hz a 16,04 s, ferme a 0,00 Hz a 16,16 s). *)
TEST 'TC-T300-BRK-040 Faute explicite : frein M3 se ferme a 10 Hz (rejeu trace 26,437 s)'
VAR
    fb : FB_Sim_TranslationBrake;
    i : INT;
END_VAR
    fb.Enable := TRUE;
    fb.ReleaseCmd := TRUE;
    fb.OpenDelay_S := 0.0;
    fb.CloseDelay_S := 0.09;
    fb.ContactDelay_S := 0.01;
    fb.CycleTime_S := 0.01;
    fb();
    ASSERT_TRUE(fb.MechanicallyOpen, 'Frein ouvert par la commande de desserrage');
    ASSERT_FALSE(fb.FaultCloseActive, 'Faute inactive par defaut');

    (* Scenario terrain : commande retiree ET variateur retournant encore 10,00 Hz. *)
    fb.ReleaseCmd := FALSE;
    fb.ActualFrequency_Hz := 10.0;
    FOR i := 1 TO 20 DO
        fb();
    END_FOR;
    ASSERT_FALSE(fb.FaultCloseActive, 'Aucune faute injectee');
    ASSERT_TRUE(fb.MechanicallyOpen, 'NOMINAL conserve : frein OUVERT a 10,00 Hz (garde 0,5 Hz)');
    ASSERT_TRUE(fb.ContactOpen, 'NOMINAL conserve : contact toujours ouvert a 10,00 Hz');

    (* Injection explicite : fermeture hors vitesse nulle, APRES le delai de faute.
       Oracle discriminateur : si le delai de faute etait ignore, la faute serait appliquee
       des le 1er scan et l'assertion ci-dessous echouerait. *)
    fb.FaultCloseWhileRunning := TRUE;
    fb.FaultCloseDelay_S := 0.5;
    FOR i := 1 TO 4 DO
        fb();
    END_FOR;
    ASSERT_FALSE(fb.FaultCloseActive, 'Faute NON appliquee avant FaultCloseDelay_S');
    ASSERT_TRUE(fb.MechanicallyOpen, 'Frein encore ouvert pendant le delai de faute');
    FOR i := 1 TO 60 DO
        fb();
    END_FOR;
    ASSERT_TRUE(fb.FaultCloseActive, 'Branche de faute appliquee apres le delai');
    ASSERT_FALSE(fb.CoilEnergized, 'Faute : bobine retombee (etat electrique coherent)');
    ASSERT_FALSE(fb.MechanicallyOpen, 'Faute : frein MECANIQUEMENT serre a 10,00 Hz');
    ASSERT_FALSE(fb.ContactOpen, 'Faute : contact frein ferme publie a 10,00 Hz');

    (* Retrait du stimulus : retour au chemin nominal, sans etat residuel. *)
    fb.FaultCloseWhileRunning := FALSE;
    fb();
    ASSERT_FALSE(fb.FaultCloseActive, 'Retrait du stimulus : faute retombee');
END_TEST

(* ---- test_fb_sim_translation_drive.st ---- *)
TEST 'TC-T300-DRV-010 Drive rampe et reponse premier ordre'
VAR
    fb : FB_Sim_TranslationDrive;
    i : INT;
END_VAR
    fb.Enable := TRUE;
    fb.FrequencyTgt_Hz := 40.0;
    fb.CycleTime_S := 0.01;
    FOR i := 1 TO 100 DO
        fb();
    END_FOR;
    ASSERT_GT(fb.FrequencyCmd_Hz, 19.7, 'Rampe 20 Hz/s apres 1 s');
    ASSERT_LT(fb.FrequencyCmd_Hz, 20.3, 'Rampe bornee apres 1 s');
    ASSERT_LT(fb.ActualFrequency_Hz, fb.FrequencyCmd_Hz, 'Retour derriere la consigne');
    ASSERT_TRUE(fb.Ready, 'Brique prete sous Enable');
END_TEST

TEST 'TC-T300-DRV-030 Charge reduit retour sans inverser la frequence'
VAR
    fb : FB_Sim_TranslationDrive;
    i : INT;
    unloaded_Hz : REAL;
END_VAR
    fb.Enable := TRUE;
    fb.FrequencyTgt_Hz := 40.0;
    fb.CycleTime_S := 0.01;
    FOR i := 1 TO 300 DO
        fb();
    END_FOR;
    unloaded_Hz := fb.ActualFrequency_Hz;
    fb.LoadAngularVelocity_RadPerS := 8.0;
    fb();
    ASSERT_LT(fb.ActualFrequency_Hz, unloaded_Hz, 'Droop charge visible au PDO');
    ASSERT_GE(fb.ActualFrequency_Hz, 0.0, 'Frequence jamais negative');
END_TEST

TEST 'TC-T300-DRV-050 Pas de 100 ms conserve le temps physique'
VAR
    fb : FB_Sim_TranslationDrive;
END_VAR
    fb.Enable := TRUE;
    fb.FrequencyTgt_Hz := 40.0;
    fb.AccelRate_HzPerS := 20.0;
    fb.CycleTime_S := 0.100;
    fb();
    ASSERT_NEAR(fb.FrequencyCmd_Hz, 2.0, 0.001,
        'A 100 ms, la rampe 20 Hz/s avance de 2 Hz');
    fb();
    ASSERT_NEAR(fb.FrequencyCmd_Hz, 4.0, 0.001,
        'Le deuxieme cycle conserve la meme duree physique');
END_TEST

(* ---- test_fb_sim_translation_dynamics.st ---- *)
(* Scenarios fonctionnels du ST reel : aucune copie du modele mecanique. *)
SETUP
VAR
    fb : FB_Sim_Translation;
    reverse : FB_Sim_Translation;
    reference : FB_Sim_Translation;
    clockProbe : FB_CycleTime;
    sensor : FB_Sim_PositionSensor;
    frequencyBefore_Hz : REAL;
    positionBefore_M : REAL;
    peakEarly_Rad : REAL;
    peakLate_Rad : REAL;
END_VAR
    fb.Enable := FALSE;
    fb();
    fb.Enable := TRUE;
    fb.ReqMaintenance := TRUE;
    fb.SpeedTgt_Pct := 40.0;
    fb.BrakeReleaseCmd := TRUE;
    fb.BrakeOpenDelayS := 0.0;
    fb.BrakeContactDelayS := 0.0;
    fb.BrakePhysicalActive := TRUE;
    fb.CartFreeActive := TRUE;
    fb.RollingFriction_Mps2 := 0.1;
    fb.SensorJitterAmplitude_M := 0.0;
END_SETUP

TEST 'M3-DYN-010 Retrait de commande a 20 Hz conserve la deceleration pilotee'
VAR
    i : INT;
END_VAR
    fb.LoadMassRatio := 0.0;
    fb.LoadReactionGain_Mps2 := 0.0;
    fb.LoadFrequencyDroopGain_Hz := 0.0;
    FOR i := 1 TO 250 DO
        fb();
    END_FOR;
    ASSERT_NEAR(fb.ActualFrequency_Hz, 20.0, 0.1, 'Regime etabli a 20 Hz');
    frequencyBefore_Hz := fb.ActualFrequency_Hz;
    positionBefore_M := fb.PositionTrue_M;
    fb.ReqMaintenance := FALSE;
    fb();
    ASSERT_GT(fb.ActualFrequency_Hz, 19.0, 'Le mot nul ne supprime pas le retour frequence');
    ASSERT_GT(fb.PositionTrue_M, positionBefore_M, 'Sens memorise pendant la deceleration');
    ASSERT_FALSE(fb.ObsCartFree, 'Pas de roue libre pendant la rampe variateur');
    FOR i := 1 TO 50 DO
        fb();
    END_FOR;
    ASSERT_LT(fb.ActualFrequency_Hz, frequencyBefore_Hz, 'Frequence decroissante');
    FOR i := 1 TO 300 DO
        fb();
    END_FOR;
    ASSERT_EQ(fb.ActualFrequency_Hz, 0.0, 'Rampe terminee');
    ASSERT_NEAR(fb.VelocityTrue_Mps, 0.0, 0.00001, 'Arret sans oscillation artificielle');
END_TEST

TEST 'M3-DYN-130 Position P1 recue initialise le chariot sans geometrie locale'
    fb.PosTremie_M := 2.0;
    fb.PosPV_M := 3.0;
    fb.PosP2_M := 5.0;
    fb.PosP1_M := 7.0;
    fb.PosMaintenance_M := 11.0;
    fb.Enable := FALSE;
    fb();
    ASSERT_NEAR(fb.PositionTrue_M, 7.0, 0.0001,
        'Repli positionne le chariot sur PosP1_M recu');
    ASSERT_TRUE(fb.PosP1, 'Repli publie P1 apres initialisation sur la position recue');
END_TEST

TEST 'M3-DYN-140 Gain recu convertit la frequence retournee en vitesse'
VAR
    i : INT;
END_VAR
    fb.PosTremie_M := 0.0;
    fb.PosPV_M := 10.0;
    fb.PosP2_M := 20.0;
    fb.PosP1_M := 30.0;
    fb.PosMaintenance_M := 40.0;
    fb.GainMetersPerHzSec := 0.03;
    fb.MaxFreq_Hz := 20.0;
    fb.Enable := FALSE;
    fb();
    fb.Enable := TRUE;
    fb.ReqMaintenance := TRUE;
    fb.SpeedTgt_Pct := 100.0;
    fb.BrakeReleaseCmd := TRUE;
    fb.BrakeOpenDelayS := 0.0;
    fb.LoadReactionGain_Mps2 := 0.0;
    FOR i := 1 TO 400 DO
        fb();
    END_FOR;
    ASSERT_NEAR(fb.ActualFrequency_Hz, 20.0, 0.05,
        'Frequence maximale recue appliquee');
    ASSERT_NEAR(fb.VelocityTrue_Mps, 0.6, 0.02,
        'Vitesse = sens x gain recu x frequence retournee');
END_TEST

TEST 'M3-DYN-100 Retour frequence electrique independant du balancement'
VAR
    drive : FB_Sim_TranslationDrive;
    i : INT;
END_VAR
    drive.Enable := TRUE;
    drive.FrequencyTgt_Hz := 20.0;
    drive.CycleTime_S := 0.01;
    FOR i := 1 TO 250 DO
        drive();
    END_FOR;
    drive.LoadAngularVelocity_RadPerS := 8.0;
    drive();
    ASSERT_NEAR(drive.ActualFrequency_Hz, drive.ElectricalFrequency_Hz, 0.00001,
        'Le retour PDO conserve la frequence electrique sous balancement');
    drive.LoadAngularVelocity_RadPerS := -8.0;
    drive();
    ASSERT_NEAR(drive.ActualFrequency_Hz, drive.ElectricalFrequency_Hz, 0.00001,
        'Pas de biais redresse par la valeur absolue du balancement');
END_TEST

TEST 'M3-DYN-110 Deceleration sans second retard sur la vitesse chariot'
VAR
    i : INT;
END_VAR
    FOR i := 1 TO 250 DO
        fb();
    END_FOR;
    fb.ReqMaintenance := FALSE;
    FOR i := 1 TO 50 DO
        fb();
    END_FOR;
    ASSERT_FALSE(fb.ObsCartFree, 'Mesure pendant la deceleration controlee');
    ASSERT_GT(fb.ActualFrequency_Hz, 5.0, 'Le variateur decelere encore');
    ASSERT_NEAR(fb.VelocityTrue_Mps, fb.ActualFrequency_Hz * 0.02, 0.001,
        'La vitesse suit le retour variateur, avec seule faible reaction mecanique');
END_TEST

TEST 'M3-DYN-120 Fin de rampe a 0.5 Hz sans supprimer consigne basse non nulle'
VAR
    drive : FB_Sim_TranslationDrive;
    i : INT;
END_VAR
    drive.Enable := TRUE;
    drive.FrequencyTgt_Hz := 20.0;
    drive.CycleTime_S := 0.01;
    FOR i := 1 TO 250 DO
        drive();
    END_FOR;
    drive.FrequencyTgt_Hz := 0.0;
    FOR i := 1 TO 120 DO
        drive();
    END_FOR;
    ASSERT_EQ(drive.ActualFrequency_Hz, 0.0, 'Fin d arret sans longue traine sous 0.5 Hz');
    drive.FrequencyTgt_Hz := 0.2;
    FOR i := 1 TO 100 DO
        drive();
    END_FOR;
    ASSERT_NEAR(drive.ActualFrequency_Hz, 0.2, 0.001,
        'Une consigne basse maintenue ne doit pas etre effacee');
END_TEST

TEST 'M3-DYN-020 Retrait brutal a 50 Hz reste limite par le variateur'
VAR
    i : INT;
END_VAR
    fb.SpeedTgt_Pct := 100.0;
    fb.LoadMassRatio := 0.0;
    fb.LoadReactionGain_Mps2 := 0.0;
    fb.LoadFrequencyDroopGain_Hz := 0.0;
    FOR i := 1 TO 400 DO
        fb();
    END_FOR;
    ASSERT_NEAR(fb.ActualFrequency_Hz, 50.0, 0.1, 'Regime etabli a 50 Hz');
    fb.ReqMaintenance := FALSE;
    positionBefore_M := fb.PositionTrue_M;
    fb();
    ASSERT_GT(fb.ActualFrequency_Hz, 49.0, 'Retour conserve apres retrait');
    ASSERT_GT(fb.PositionTrue_M, positionBefore_M, 'Pas de gel de position au retrait');
    ASSERT_FALSE(fb.ObsCartFree, 'Variateur encore en deceleration');
    FOR i := 1 TO 400 DO
        fb();
    END_FOR;
    ASSERT_EQ(fb.ActualFrequency_Hz, 0.0, 'Frequence finalement nulle');
    ASSERT_NEAR(fb.VelocityTrue_Mps, 0.0, 0.00001, 'Arret final');
    ASSERT_FALSE(fb.HardStopMaintenanceActive, 'Arret observe hors butee');
END_TEST

TEST 'M3-DYN-030 Frottement seul a 100 ms sans inversion dans les deux sens'
    fb.SpeedTgt_Pct := 0.4;
    fb.DriveTimeConstantS := 0.0;
    fb.LoadMassRatio := 0.0;
    fb.LoadReactionGain_Mps2 := 0.0;
    fb.LoadFrequencyDroopGain_Hz := 0.0;
    fb();
    reverse(Enable := TRUE, ReqTremie := TRUE, SpeedTgt_Pct := 0.4,
        BrakeReleaseCmd := TRUE, BrakeOpenDelayS := 0.0, DriveTimeConstantS := 0.0,
        CartFreeActive := TRUE, RollingFriction_Mps2 := 0.1, LoadMassRatio := 0.0,
        LoadReactionGain_Mps2 := 0.0, LoadFrequencyDroopGain_Hz := 0.0);
    ASSERT_NEAR(fb.VelocityTrue_Mps, 0.004, 0.00001, 'Petite vitesse positive initiale');
    ASSERT_NEAR(reverse.VelocityTrue_Mps, -0.004, 0.00001, 'Petite vitesse negative initiale');
    clockProbe();
    fb.ReqMaintenance := FALSE;
    reverse.ReqTremie := FALSE;
    ADVANCE_TIME(100000000);
    clockProbe();
    ASSERT_NEAR(clockProbe.CycleTimeS, 0.1, 0.00001, 'Pas reel de 100 ms');
    fb();
    reverse();
    ASSERT_EQ(fb.VelocityTrue_Mps, 0.0, 'Frottement arrete le sens positif sans inversion');
    ASSERT_EQ(reverse.VelocityTrue_Mps, 0.0, 'Frottement arrete le sens negatif sans inversion');
    ASSERT_TRUE(fb.ObsCartFree, 'Le calcul libre est effectivement exerce');
    ADVANCE_TIME(100000000);
    fb();
    reverse();
    ASSERT_EQ(fb.VelocityTrue_Mps, 0.0, 'Pas de redemarrage numerique positif');
    ASSERT_EQ(reverse.VelocityTrue_Mps, 0.0, 'Pas de redemarrage numerique negatif');
END_TEST

TEST 'M3-DYN-040 Frottement seul a 10 ms sans inversion dans les deux sens'
    fb.SpeedTgt_Pct := 0.04;
    fb.DriveTimeConstantS := 0.0;
    fb.LoadMassRatio := 0.0;
    fb.LoadReactionGain_Mps2 := 0.0;
    fb.LoadFrequencyDroopGain_Hz := 0.0;
    fb();
    reverse(Enable := TRUE, ReqTremie := TRUE, SpeedTgt_Pct := 0.04,
        BrakeReleaseCmd := TRUE, BrakeOpenDelayS := 0.0, DriveTimeConstantS := 0.0,
        CartFreeActive := TRUE, RollingFriction_Mps2 := 0.1, LoadMassRatio := 0.0,
        LoadReactionGain_Mps2 := 0.0, LoadFrequencyDroopGain_Hz := 0.0);
    clockProbe();
    fb.ReqMaintenance := FALSE;
    reverse.ReqTremie := FALSE;
    ADVANCE_TIME(10000000);
    clockProbe();
    ASSERT_NEAR(clockProbe.CycleTimeS, 0.01, 0.00001, 'Pas reel de 10 ms');
    fb();
    reverse();
    ASSERT_EQ(fb.VelocityTrue_Mps, 0.0, 'Immobilite positive conservee');
    ASSERT_EQ(reverse.VelocityTrue_Mps, 0.0, 'Immobilite negative conservee');
END_TEST

TEST 'M3-DYN-050 Adherence au repos et au seuil puis depart sous poussee'
    (* Seuil explicite du scenario historique ; ne calibre pas le banc. *)
    fb.StaticFriction_Mps2 := 0.1;
    fb.ReqMaintenance := FALSE;
    fb.LoadMassRatio := 0.0;
    fb.Slope_Mps2 := 0.05;
    fb();
    ASSERT_EQ(fb.VelocityTrue_Mps, 0.0, 'Poussee sous le frottement : immobile');
    fb.Slope_Mps2 := 0.1;
    fb();
    ASSERT_EQ(fb.VelocityTrue_Mps, 0.0, 'Poussee au seuil : immobile');
    fb.Slope_Mps2 := 0.2;
    fb();
    ASSERT_GT(fb.VelocityTrue_Mps, 0.0, 'Poussee suffisante : depart physique');
END_TEST

TEST 'M3-DYN-051 Pente seule au repos respecte le seuil statique courant'
VAR
    i : INT;
END_VAR
    fb.ReqMaintenance := FALSE;
    fb.LoadMassRatio := 0.0;
    fb.LoadReactionGain_Mps2 := 0.0;
    fb.StaticFriction_Mps2 := 0.35;
    fb.RollingFriction_Mps2 := 0.30;
    fb.Slope_Mps2 := 0.20;
    positionBefore_M := fb.PositionTrue_M;
    FOR i := 1 TO 100 DO
        fb();
    END_FOR;
    ASSERT_EQ(fb.VelocityTrue_Mps, 0.0, 'Pente sous adhesion : aucun depart');
    fb.Slope_Mps2 := 0.35;
    fb();
    ASSERT_EQ(fb.VelocityTrue_Mps, 0.0, 'Au seuil statique : aucun depart');
    fb.Slope_Mps2 := 0.60;
    fb();
    ASSERT_GT(fb.VelocityTrue_Mps, 0.0, 'Pente au-dessus adhesion : depart');
    ASSERT_TRUE(fb.ObsCartFree, 'Frein ouvert sans couple variateur');
END_TEST

TEST 'M3-DYN-052 Frein ferme retient une pente puis ouverture autorise derive'
VAR
    i : INT;
END_VAR
    fb.ReqMaintenance := FALSE;
    fb.BrakeReleaseCmd := FALSE;
    fb.LoadMassRatio := 0.0;
    fb.LoadReactionGain_Mps2 := 0.0;
    fb.StaticFriction_Mps2 := 0.35;
    fb.RollingFriction_Mps2 := 0.30;
    fb.Slope_Mps2 := -0.60;
    fb();
    positionBefore_M := fb.PositionTrue_M;
    FOR i := 1 TO 100 DO
        fb();
    END_FOR;
    ASSERT_EQ(fb.PositionTrue_M, positionBefore_M, 'Frein ferme : pente sans mouvement');
    ASSERT_FALSE(fb.ObsCartFree, 'Pas de regime libre frein ferme');
    fb.BrakeReleaseCmd := TRUE;
    fb();
    ASSERT_TRUE(fb.ObsCartFree, 'Relachement frein : regime libre');
    ASSERT_LT(fb.PositionTrue_M, positionBefore_M, 'Pente negative : mouvement vers Tremie');
    fb.BrakeReleaseCmd := FALSE;
    FOR i := 1 TO 100 DO
        fb();
    END_FOR;
    ASSERT_FALSE(fb.BrakeMechanicallyOpen, 'Frein referme');
    ASSERT_EQ(fb.VelocityTrue_Mps, 0.0, 'Frein arrete la derive');
END_TEST

TEST 'M3-DYN-060 Poussee opposee suffisante autorise une vraie inversion'
    fb.SpeedTgt_Pct := 0.4;
    fb.DriveTimeConstantS := 0.0;
    fb.LoadMassRatio := 0.0;
    fb.LoadReactionGain_Mps2 := 0.0;
    fb.LoadFrequencyDroopGain_Hz := 0.0;
    fb();
    ASSERT_GT(fb.VelocityTrue_Mps, 0.0, 'Vitesse initiale positive');
    fb.ReqMaintenance := FALSE;
    (* Force superieure au seuil statique 0.35 : inversion physiquement autorisee. *)
    fb.Slope_Mps2 := -0.6;
    ADVANCE_TIME(100000000);
    fb();
    ASSERT_LT(fb.VelocityTrue_Mps, 0.0, 'La correction ne bloque pas une vraie inversion');
END_TEST

TEST 'M3-DYN-070 Frein ferme en mouvement suit la bobine sans attendre les Hz'
VAR
    i : INT;
END_VAR
    FOR i := 1 TO 250 DO
        fb();
    END_FOR;
    ASSERT_GT(fb.VelocityTrue_Mps, 0.3, 'Chariot initialement en mouvement');
    fb.BrakeReleaseCmd := FALSE;
    fb();
    ASSERT_FALSE(fb.BrakeCoilEnergized, 'Coupure bobine immediate');
    ASSERT_TRUE(fb.BrakeMechanicallyOpen, 'Delai mecanique conserve');
    FOR i := 1 TO 60 DO
        fb();
    END_FOR;
    ASSERT_FALSE(fb.BrakeMechanicallyOpen, 'Frein serre malgre frequence non nulle');
    ASSERT_FALSE(fb.BrakeContactOpen, 'Retour frein ferme');
    ASSERT_GT(fb.ActualFrequency_Hz, 10.0, 'La sortie variateur est encore non nulle');
    ASSERT_EQ(fb.VelocityTrue_Mps, 0.0, 'Frein immobilise le chariot');
    ASSERT_EQ(fb.ObsBrakeClosedMovingCount, 1, 'Fermeture en mouvement observable');
END_TEST

TEST 'M3-DYN-080 Balancement conserve secondaire sous controle puis amorti'
VAR
    i : INT;
END_VAR
    reference.Enable := TRUE;
    reference.ReqMaintenance := TRUE;
    reference.SpeedTgt_Pct := 40.0;
    reference.BrakeReleaseCmd := TRUE;
    reference.BrakeOpenDelayS := 0.0;
    reference.SuspendedLoadLength_M := 0.0;
    FOR i := 1 TO 300 DO
        fb();
        reference();
    END_FOR;
    ASSERT_TRUE(ABS(fb.LoadAngle_Rad) > 0.0001, 'Balancement present');
    ASSERT_LT(ABS(fb.PositionTrue_M - reference.PositionTrue_M), 0.05,
        'Contribution secondaire dans ce scenario fixe, sans plafonnement de distance');
    ASSERT_FALSE(fb.ObsCartFree, 'Comparaison effectuee sous controle variateur');
    fb.ReqMaintenance := FALSE;
    fb.BrakeReleaseCmd := FALSE;
    FOR i := 1 TO 800 DO
        fb();
        IF i <= 100 THEN
            peakEarly_Rad := MAX(peakEarly_Rad, ABS(fb.LoadAngle_Rad));
        END_IF;
        IF i > 700 THEN
            peakLate_Rad := MAX(peakLate_Rad, ABS(fb.LoadAngle_Rad));
        END_IF;
    END_FOR;
    ASSERT_GT(peakEarly_Rad, 0.001, 'Pendule excite par le freinage');
    ASSERT_LT(peakLate_Rad, peakEarly_Rad, 'Oscillations amorties');
    ASSERT_EQ(fb.VelocityTrue_Mps, 0.0, 'Pendule ne deplace pas le frein serre');
END_TEST

TEST 'M3-DYN-090 Came spatiale vue perdue retrouvee stable sans blip ajoute'
    sensor(Enable := TRUE, Position_M := 0.2, Threshold_M := 0.0,
        CamDropoutActive := TRUE, CamDropoutStart_M := 0.02, CamDropoutWidth_M := 0.04,
        ElectricalDelayS := 0.0, IntermittenceActive := FALSE, BlipTransitions := 0);
    ASSERT_FALSE(sensor.ElectricalOutput, 'Avant la detection');
    sensor(Position_M := -0.03);
    ASSERT_TRUE(sensor.ElectricalOutput, 'Cible vue');
    sensor(Position_M := -0.06);
    ASSERT_FALSE(sensor.ElectricalOutput, 'Interruption de cible');
    sensor(Position_M := -0.10);
    ASSERT_TRUE(sensor.ElectricalOutput, 'Cible retrouvee');
    sensor();
    ASSERT_TRUE(sensor.ElectricalOutput, 'Etat stable sans intermittence temporelle');
    sensor(Position_M := -0.06);
    ASSERT_FALSE(sensor.ElectricalOutput, 'Zone de perte aussi au retour');
    sensor(Position_M := -0.02);
    ASSERT_TRUE(sensor.ElectricalOutput, 'Cible retrouvee au retour');
    sensor(Position_M := 0.03);
    ASSERT_FALSE(sensor.ElectricalOutput, 'Sortie de cible');
END_TEST

(* ---- test_fb_sim_translation_t417_boundary.st ---- *)
(* T417 investigation : vitesse initiale opposee a une force inferieure au seuil
   statique. Apres passage a zero, cette force ne peut pas redemarrer le chariot.
   Parametres synthetiques explicites, aucune calibration terrain. *)
SETUP
VAR
    fb : FB_Sim_Translation;
    reverse : FB_Sim_Translation;
END_VAR
    fb(Enable := FALSE);
    reverse(Enable := FALSE);
    fb(Enable := TRUE, ReqMaintenance := TRUE, SpeedTgt_Pct := 0.4,
        BrakeReleaseCmd := TRUE, BrakeOpenDelayS := 0.0, DriveTimeConstantS := 0.0,
        CartFreeActive := TRUE, RollingFriction_Mps2 := 0.1, StaticFriction_Mps2 := 0.35,
        LoadMassRatio := 0.0, LoadReactionGain_Mps2 := 0.0, SensorJitterAmplitude_M := 0.0);
    reverse(Enable := TRUE, ReqTremie := TRUE, SpeedTgt_Pct := 0.4,
        BrakeReleaseCmd := TRUE, BrakeOpenDelayS := 0.0, DriveTimeConstantS := 0.0,
        CartFreeActive := TRUE, RollingFriction_Mps2 := 0.1, StaticFriction_Mps2 := 0.35,
        LoadMassRatio := 0.0, LoadReactionGain_Mps2 := 0.0, SensorJitterAmplitude_M := 0.0);
END_SETUP

TEST 'T417-BOUND-010 Force opposee sous seuil statique ne redemarre pas apres zero'
    ASSERT_NEAR(fb.VelocityTrue_Mps, 0.004, 0.00001, 'Vitesse initiale positive');
    fb.ReqMaintenance := FALSE;
    fb.Slope_Mps2 := -0.2;
    ADVANCE_TIME(100000000);
    fb();
    ASSERT_TRUE(fb.ObsCartFree, 'Branche libre exercee');
    ASSERT_EQ(fb.VelocityTrue_Mps, 0.0, 'Arret puis adherence : force 0.2 inferieure au seuil 0.35');
END_TEST

TEST 'T417-BOUND-040 Frottement banc 0.30 et pas 100 ms respectent adherence'
    fb.SpeedTgt_Pct := 0.2;
    fb.RollingFriction_Mps2 := 0.30;
    fb();
    ASSERT_NEAR(fb.VelocityTrue_Mps, 0.002, 0.00001, 'Vitesse avant arret');
    fb.ReqMaintenance := FALSE;
    fb.Slope_Mps2 := -0.34;
    ADVANCE_TIME(100000000);
    fb();
    ASSERT_TRUE(fb.ObsCartFree, 'Branche libre exercee');
    ASSERT_EQ(fb.VelocityTrue_Mps, 0.0, 'Force 0.34 sous seuil 0.35 : adherence apres zero');
END_TEST

TEST 'T417-BOUND-050 Meme scenario avec pas 20 ms'
    fb.SpeedTgt_Pct := 0.2;
    fb.RollingFriction_Mps2 := 0.30;
    fb();
    ASSERT_NEAR(fb.VelocityTrue_Mps, 0.002, 0.00001, 'Vitesse avant arret');
    fb.ReqMaintenance := FALSE;
    fb.Slope_Mps2 := -0.34;
    ADVANCE_TIME(20000000);
    fb();
    ASSERT_TRUE(fb.ObsCartFree, 'Branche libre exercee');
    ASSERT_EQ(fb.VelocityTrue_Mps, 0.0, 'Meme verdict adherence au pas 20 ms');
END_TEST

TEST 'T417-BOUND-020 Meme adherence dans le sens negatif'
    ASSERT_NEAR(reverse.VelocityTrue_Mps, -0.004, 0.00001, 'Vitesse initiale negative');
    reverse.ReqTremie := FALSE;
    reverse.Slope_Mps2 := 0.2;
    ADVANCE_TIME(100000000);
    reverse();
    ASSERT_TRUE(reverse.ObsCartFree, 'Branche libre exercee');
    ASSERT_EQ(reverse.VelocityTrue_Mps, 0.0, 'Arret puis adherence symetrique');
END_TEST

TEST 'T417-BOUND-030 Une force au dessus du seuil permet inversion'
    fb.ReqMaintenance := FALSE;
    fb.Slope_Mps2 := -0.6;
    ADVANCE_TIME(100000000);
    fb();
    ASSERT_TRUE(fb.ObsCartFree, 'Branche libre exercee');
    ASSERT_LT(fb.VelocityTrue_Mps, 0.0, 'Force 0.6 superieure au seuil 0.35 : inversion autorisee');
END_TEST

TEST 'T417-BOUND-060 Force exactement au seuil statique reste collee au croisement'
    fb.SpeedTgt_Pct := 0.4;
    fb.RollingFriction_Mps2 := 0.1;
    fb.StaticFriction_Mps2 := 0.35;
    fb();
    ASSERT_NEAR(fb.VelocityTrue_Mps, 0.004, 0.00001, 'Vitesse initiale positive');
    fb.ReqMaintenance := FALSE;
    fb.Slope_Mps2 := -0.35;
    ADVANCE_TIME(100000000);
    fb();
    ASSERT_EQ(fb.VelocityTrue_Mps, 0.0, 'Comparaison inclusive : egalite = adhesion');
END_TEST

TEST 'T417-BOUND-070 Prediction exactement nulle et force supra seuil'
    fb.SpeedTgt_Pct := 0.4;
    fb.RollingFriction_Mps2 := 0.1;
    fb.StaticFriction_Mps2 := 0.35;
    fb();
    ASSERT_NEAR(fb.VelocityTrue_Mps, 0.004, 0.00001, 'Vitesse initiale positive');
    fb.ReqMaintenance := FALSE;
    fb.Slope_Mps2 := -0.04;
    ADVANCE_TIME(100000000);
    fb();
    ASSERT_EQ(fb.VelocityTrue_Mps, 0.0, 'Prediction nulle garde le mouvement pour ce scan');
END_TEST

TEST 'T417-BOUND-080 Seuil de vitesse 0.001 distingue repos et mouvement'
    fb.SpeedTgt_Pct := 0.1;
    fb.RollingFriction_Mps2 := 0.0;
    fb.StaticFriction_Mps2 := 0.35;
    fb.Slope_Mps2 := 0.0;
    fb();
    ASSERT_NEAR(fb.VelocityTrue_Mps, 0.001, 0.00001, 'Vitesse au seuil');
    fb.SpeedTgt_Pct := 0.08;
    fb();
    ASSERT_NEAR(fb.VelocityTrue_Mps, 0.0008, 0.00001, 'Vitesse sous seuil');
END_TEST
